(* IEC 61131-3 sources: plc-vscode/tests/st/all/trust-platform/examples/OSCAT/tunnel_oven_strategy_observer/oop/src, 3 files *)

(* ---- Main.st ---- *)
(* Pattern role: IOvenProfile is the contract boundary for the Strategy and Observer example. *)
INTERFACE IOvenProfile
    PROPERTY ProfileId : INT
    GET
    END_GET
    END_PROPERTY

    METHOD HeatCommand : REAL
    VAR_INPUT
        ZoneTemp : REAL;
    END_VAR
    END_METHOD

    METHOD ConveyorSpeed : REAL
    END_METHOD
END_INTERFACE

(* Pattern role: IOvenEventSubscriber is the contract boundary for the Strategy and Observer example. *)
INTERFACE IOvenEventSubscriber
    METHOD OnOvenEvent
    VAR_INPUT
        EventClass : BYTE;
        EventCode : WORD;
        ProfileId : INT;
    END_VAR
    END_METHOD
END_INTERFACE

(* Pattern role: BreadProfile is a concrete implementation in the Strategy and Observer example. *)
FUNCTION_BLOCK BreadProfile IMPLEMENTS IOvenProfile
VAR
    Filter : Pt1Filter;
END_VAR

METHOD PUBLIC Initialize
Filter.Initialize();
Filter.Configure(TimeConstant := T#3s, Gain := REAL#1.0);
END_METHOD

METHOD PUBLIC HeatCommand : REAL
VAR_INPUT
    ZoneTemp : REAL;
END_VAR
HeatCommand := LIMIT(REAL#0.0, (REAL#185.0 - Filter.Update(Sample := ZoneTemp)) * REAL#1.5, REAL#100.0);
END_METHOD

METHOD PUBLIC ConveyorSpeed : REAL
ConveyorSpeed := REAL#35.0;
END_METHOD

PUBLIC PROPERTY ProfileId : INT
GET
    ProfileId := INT#1;
END_GET
END_PROPERTY
END_FUNCTION_BLOCK

(* Pattern role: PizzaProfile is a concrete implementation in the Strategy and Observer example. *)
FUNCTION_BLOCK PizzaProfile IMPLEMENTS IOvenProfile
VAR
    Filter : Pt1Filter;
END_VAR

METHOD PUBLIC Initialize
Filter.Initialize();
Filter.Configure(TimeConstant := T#1s, Gain := REAL#1.0);
END_METHOD

METHOD PUBLIC HeatCommand : REAL
VAR_INPUT
    ZoneTemp : REAL;
END_VAR
HeatCommand := LIMIT(REAL#0.0, (REAL#235.0 - Filter.Update(Sample := ZoneTemp)) * REAL#2.0, REAL#100.0);
END_METHOD

METHOD PUBLIC ConveyorSpeed : REAL
ConveyorSpeed := REAL#55.0;
END_METHOD

PUBLIC PROPERTY ProfileId : INT
GET
    ProfileId := INT#2;
END_GET
END_PROPERTY
END_FUNCTION_BLOCK

(* Pattern role: OvenHistorianSubscriber is a concrete implementation in the Strategy and Observer example. *)
FUNCTION_BLOCK OvenHistorianSubscriber IMPLEMENTS IOvenEventSubscriber
VAR
    EventCountValue : INT;
END_VAR

METHOD PUBLIC OnOvenEvent
VAR_INPUT
    EventClass : BYTE;
    EventCode : WORD;
    ProfileId : INT;
END_VAR
EventCountValue := EventCountValue + INT#1;
END_METHOD

PUBLIC PROPERTY EventCount : INT
GET
    EventCount := EventCountValue;
END_GET
END_PROPERTY
END_FUNCTION_BLOCK

(* Pattern role: OvenMqttSubscriber is a concrete implementation in the Strategy and Observer example. *)
FUNCTION_BLOCK OvenMqttSubscriber IMPLEMENTS IOvenEventSubscriber
VAR
    PublishReadyValue : BOOL;
END_VAR

METHOD PUBLIC OnOvenEvent
VAR_INPUT
    EventClass : BYTE;
    EventCode : WORD;
    ProfileId : INT;
END_VAR
PublishReadyValue := TRUE;
END_METHOD

PUBLIC PROPERTY PublishReady : BOOL
GET
    PublishReady := PublishReadyValue;
END_GET
END_PROPERTY
END_FUNCTION_BLOCK

(* Composition role: OvenEventBus owns the collaborating objects used by this Strategy and Observer example. *)
FUNCTION_BLOCK OvenEventBus
VAR
    Historian : IOvenEventSubscriber;
    Mqtt : IOvenEventSubscriber;
END_VAR

METHOD PUBLIC Subscribe
VAR_INPUT
    HistorianSub : IOvenEventSubscriber;
    MqttSub : IOvenEventSubscriber;
END_VAR
Historian := HistorianSub;
Mqtt := MqttSub;
END_METHOD

METHOD PUBLIC Publish
VAR_INPUT
    EventClass : BYTE;
    EventCode : WORD;
    ProfileId : INT;
END_VAR
Historian.OnOvenEvent(EventClass := EventClass, EventCode := EventCode, ProfileId := ProfileId);
Mqtt.OnOvenEvent(EventClass := EventClass, EventCode := EventCode, ProfileId := ProfileId);
END_METHOD
END_FUNCTION_BLOCK

(* Composition role: TunnelOvenController owns the collaborating objects used by this Strategy and Observer example. *)
FUNCTION_BLOCK TunnelOvenController
VAR
    Bread : BreadProfile;
    Pizza : PizzaProfile;
    ActiveProfile : IOvenProfile;
    Bus : OvenEventBus;
    Historian : OvenHistorianSubscriber;
    Mqtt : OvenMqttSubscriber;
    ActiveProfileIdValue : INT;
    ZoneHeatCommandValue : REAL;
    ConveyorSpeedValue : REAL;
END_VAR

METHOD PUBLIC Initialize
Bread.Initialize();
Pizza.Initialize();
Bus.Subscribe(HistorianSub := Historian, MqttSub := Mqtt);
ActiveProfile := Bread;
END_METHOD

METHOD PUBLIC SelectProfile
VAR_INPUT
    ProductId : INT;
END_VAR
IF ProductId = INT#2 THEN
    ActiveProfile := Pizza;
ELSE
    ActiveProfile := Bread;
END_IF;
ActiveProfileIdValue := ActiveProfile.ProfileId;
END_METHOD

METHOD PUBLIC Update : REAL
VAR_INPUT
    ProductId : INT;
    ZoneTemp : REAL;
    Overtemp : BOOL;
END_VAR
SelectProfile(ProductId := ProductId);
ZoneHeatCommandValue := ActiveProfile.HeatCommand(ZoneTemp := ZoneTemp);
ConveyorSpeedValue := ActiveProfile.ConveyorSpeed();
IF Overtemp THEN
    ZoneHeatCommandValue := REAL#0.0;
    Bus.Publish(EventClass := BYTE#3, EventCode := WORD#16#A601, ProfileId := ActiveProfile.ProfileId);
END_IF;
Update := ZoneHeatCommandValue;
END_METHOD

PUBLIC PROPERTY ActiveProfileId : INT
GET
    ActiveProfileId := ActiveProfileIdValue;
END_GET
END_PROPERTY

PUBLIC PROPERTY ZoneHeatCommand : REAL
GET
    ZoneHeatCommand := ZoneHeatCommandValue;
END_GET
END_PROPERTY

PUBLIC PROPERTY ConveyorSpeed : REAL
GET
    ConveyorSpeed := ConveyorSpeedValue;
END_GET
END_PROPERTY

PUBLIC PROPERTY QualityEventCount : INT
GET
    QualityEventCount := Historian.EventCount;
END_GET
END_PROPERTY

PUBLIC PROPERTY MqttPublishReady : BOOL
GET
    MqttPublishReady := Mqtt.PublishReady;
END_GET
END_PROPERTY
END_FUNCTION_BLOCK

(* Scan role: Main wires the example objects and exposes the PLC call path under test. *)
PROGRAM Main
VAR
    Oven : TunnelOvenController;
    ProductId : INT;
    ZoneTempRaw : INT;
    OvertempInput : BOOL;
    HeatCommandRaw : INT;
    ConveyorSpeedRaw : INT;
    AlarmOut : BOOL;
END_VAR

Oven.Initialize();
HeatCommandRaw := REAL_TO_INT(Oven.Update(ProductId := ProductId, ZoneTemp := INT_TO_REAL(ZoneTempRaw), Overtemp := OvertempInput));
ConveyorSpeedRaw := REAL_TO_INT(Oven.ConveyorSpeed);
AlarmOut := Oven.QualityEventCount > INT#0;
END_PROGRAM

(* ---- Configuration.st ---- *)
CONFIGURATION TunnelOvenStrategyObserverOopConfiguration
RESOURCE Cpu0 ON PLC
    TASK MainTask (INTERVAL := T#100ms, PRIORITY := 1);
    PROGRAM Oven WITH MainTask : Main;
END_RESOURCE
VAR_CONFIG
    Oven.ProductId AT %IW0 : INT;
    Oven.ZoneTempRaw AT %IW2 : INT;
    Oven.OvertempInput AT %IX0.0 : BOOL;
    Oven.HeatCommandRaw AT %QW0 : INT;
    Oven.ConveyorSpeedRaw AT %QW2 : INT;
    Oven.AlarmOut AT %QX0.0 : BOOL;
END_VAR
END_CONFIGURATION

(* ---- Tests.st ---- *)
TEST_PROGRAM OvenStrategiesProduceDifferentCommands
VAR
    Oven : TunnelOvenController;
    BreadHeat : REAL;
    PizzaHeat : REAL;
END_VAR

Oven.Initialize();
BreadHeat := Oven.Update(ProductId := INT#1, ZoneTemp := REAL#180.0, Overtemp := FALSE);
ASSERT_EQUAL(EXPECTED := INT#1, ACTUAL := Oven.ActiveProfileId);
PizzaHeat := Oven.Update(ProductId := INT#2, ZoneTemp := REAL#180.0, Overtemp := FALSE);
ASSERT_EQUAL(EXPECTED := INT#2, ACTUAL := Oven.ActiveProfileId);
ASSERT_TRUE(IN := PizzaHeat > BreadHeat);
ASSERT_NEAR(EXPECTED := REAL#55.0, ACTUAL := Oven.ConveyorSpeed, DELTA := REAL#0.001);
END_TEST_PROGRAM

TEST_PROGRAM OvenObserverPublishesOvertempEvent
VAR
    Oven : TunnelOvenController;
    Heat : REAL;
END_VAR

Oven.Initialize();
Heat := Oven.Update(ProductId := INT#2, ZoneTemp := REAL#260.0, Overtemp := TRUE);
ASSERT_NEAR(EXPECTED := REAL#0.0, ACTUAL := Heat, DELTA := REAL#0.001);
ASSERT_EQUAL(EXPECTED := INT#1, ACTUAL := Oven.QualityEventCount);
ASSERT_TRUE(IN := Oven.MqttPublishReady);
END_TEST_PROGRAM

(* Multi-event observer + strategy test: drives the same oven through
   normal -> overtemp -> recovered with a profile switch. Catches bugs
   where QualityEventCount stops growing after the first event or
   where the strategy slot fails to re-evaluate when ProductId changes
   after an overtemp recovery. *)
TEST_PROGRAM OvenAccumulatesEventsAndSwitchesProfileAcrossScans
VAR
    Oven : TunnelOvenController;
    InitialEvents : INT;
END_VAR

Oven.Initialize();

(* Scan 1: normal pizza bake *)
Oven.Update(ProductId := INT#2, ZoneTemp := REAL#180.0, Overtemp := FALSE);
InitialEvents := Oven.QualityEventCount;

(* Scan 2: overtemp event - count must grow *)
Oven.Update(ProductId := INT#2, ZoneTemp := REAL#260.0, Overtemp := TRUE);
ASSERT_TRUE(IN := Oven.QualityEventCount > InitialEvents);

(* Scan 3: recovered, switched to bread profile *)
Oven.Update(ProductId := INT#1, ZoneTemp := REAL#180.0, Overtemp := FALSE);
ASSERT_EQUAL(EXPECTED := INT#1, ACTUAL := Oven.ActiveProfileId);
END_TEST_PROGRAM

(* Multi-call regression: every overtemp on a single scan increments the
   historian counter exactly once. Catches bugs where the observer fires
   twice (e.g., once per profile member access) or zero times (e.g.,
   if the bus publishes to a stale subscriber slot). *)
TEST_PROGRAM OvenObserverIncrementsExactlyOncePerOvertempScan
VAR
    Oven : TunnelOvenController;
    I : INT;
    ExpectedCount : INT;
END_VAR

Oven.Initialize();
ExpectedCount := INT#0;
FOR I := 1 TO 5 DO
    Oven.Update(ProductId := INT#2, ZoneTemp := REAL#260.0, Overtemp := TRUE);
    ExpectedCount := ExpectedCount + INT#1;
    ASSERT_EQUAL(EXPECTED := ExpectedCount, ACTUAL := Oven.QualityEventCount);
END_FOR;
END_TEST_PROGRAM

(* Boundary test: well below setpoint, the LIMIT clamps the bread
   heat command to 100. (Pt1Filter is wall-clock based so chasing high
   inputs from a cold first sample is not stable in microsecond test
   cycles; we only check the cold-clamp here.) *)
TEST_PROGRAM OvenBreadProfileColdClampsHeatCommandHigh
VAR
    Oven : TunnelOvenController;
    Heat : REAL;
END_VAR

Oven.Initialize();
Heat := Oven.Update(ProductId := INT#1, ZoneTemp := REAL#20.0, Overtemp := FALSE);
ASSERT_NEAR(EXPECTED := REAL#100.0, ACTUAL := Heat, DELTA := REAL#0.5);
END_TEST_PROGRAM

(* Per-FB isolation: directly drive a PizzaProfile object and verify it
   reports profile id 2 and conveyor speed 55 without a controller. *)
TEST_PROGRAM OvenPizzaProfileReportsExpectedConveyorAndId
VAR
    Pizza : PizzaProfile;
    Speed : REAL;
END_VAR

Pizza.Initialize();
ASSERT_EQUAL(EXPECTED := INT#2, ACTUAL := Pizza.ProfileId);
Speed := Pizza.ConveyorSpeed();
ASSERT_NEAR(EXPECTED := REAL#55.0, ACTUAL := Speed, DELTA := REAL#0.001);
END_TEST_PROGRAM

(* Per-FB isolation: drive an OvenHistorianSubscriber on its own and
   confirm that EventCount accumulates one per OnOvenEvent call. *)
TEST_PROGRAM OvenHistorianSubscriberCountsAllEvents
VAR
    Sub : OvenHistorianSubscriber;
END_VAR

Sub.OnOvenEvent(EventClass := BYTE#3, EventCode := WORD#16#A601, ProfileId := INT#1);
Sub.OnOvenEvent(EventClass := BYTE#3, EventCode := WORD#16#A601, ProfileId := INT#2);
Sub.OnOvenEvent(EventClass := BYTE#1, EventCode := WORD#16#B001, ProfileId := INT#2);
ASSERT_EQUAL(EXPECTED := INT#3, ACTUAL := Sub.EventCount);
END_TEST_PROGRAM

(* Edge input: ProductId outside {1, 2} must default to bread (id 1)
   so a stale or wild input never selects an undefined strategy. *)
TEST_PROGRAM OvenUnknownProductIdDefaultsToBread
VAR
    Oven : TunnelOvenController;
END_VAR

Oven.Initialize();
Oven.Update(ProductId := INT#42, ZoneTemp := REAL#180.0, Overtemp := FALSE);
ASSERT_EQUAL(EXPECTED := INT#1, ACTUAL := Oven.ActiveProfileId);
ASSERT_NEAR(EXPECTED := REAL#35.0, ACTUAL := Oven.ConveyorSpeed, DELTA := REAL#0.001);
Oven.Update(ProductId := INT#-1, ZoneTemp := REAL#180.0, Overtemp := FALSE);
ASSERT_EQUAL(EXPECTED := INT#1, ACTUAL := Oven.ActiveProfileId);
END_TEST_PROGRAM
